VAR_GLOBAL
    bUpperButton AT %I* : BOOL;
    bLowerButton AT %I* : BOOL;
    bOuterSpotsRelay AT %Q* : BOOL;
    bMiddleSpotRelay AT %Q* : BOOL;
END_VAR

(* stored: Version 1.1.0.1
   GVL GVL_HallIO: Id {7ba4e0f5-2971-47d5-a58a-b437d57a7d77} *)
